Fanuc KAREL source: kt00646.KL

-- PROVISIONAL review KL for V770-1; original PC SHA256 6738c83e93aeb60af3fe00269f1459456c9c09c1b004dfffbdb615573fa0ea32
-- Incomplete behavior may be omitted. Consult companion uncertainty JSON. Do not deploy.
PROGRAM KT00646
%NOLOCKGROUP
VAR
  OUT : INTEGER
-- UNRESOLVED_DECL H1 type=002017
-- UNRESOLVED_DECL H2 type=002017
BEGIN
  -- UNRESOLVED_PC offsets 5-19; opcodes 2E,22,9D,33,B4
  -- UNRESOLVED_PC offsets 24-38; opcodes 2E,22,9D,33,B4
  -- UNRESOLVED_PC offsets 43-57; opcodes 2E,22,9D,33,B4
  -- UNRESOLVED_PC offsets 62-76; opcodes 2E,22,9D,33,B4
  -- UNRESOLVED_PC offsets 81-96; opcodes 22,9D,33,B3,23
  -- UNRESOLVED_PC offsets 101-105; opcodes 7F
END KT00646
